Fanuc KAREL source: kb00111.KL

-- PROVISIONAL review KL for V770-1; original PC SHA256 cd52c107ac11bb60356b7f60936e3e6edd0103f86a375c0b045788f3049409d8
-- Incomplete behavior may be omitted. Consult companion uncertainty JSON. Do not deploy.
PROGRAM KB00111
%NOLOCKGROUP
BEGIN
  -- UNRESOLVED_PC offsets 5-21; opcodes 27,22,31,23
  -- UNRESOLVED_PC offsets 26-30; opcodes 7F
END KB00111
